TYPE "ST_DeclarationParCfg"
VERSION : 0.1
   STRUCT
      SchemaVersion : UInt := 3;
      Timeout : Time := T#2S;
   END_STRUCT;

END_TYPE

